Fanuc KAREL source: KT00067.KL

PROGRAM KT00067
%NOLOCKGROUP
VAR
  I1: INTEGER
  R2: REAL
  OUT: INTEGER
BEGIN
  I1 = 2
    R2 = 3.0
  OUT = I1 * R2
END KT00067
